(* Schneider Machine Expert - Basic project Projeto Charpy 3 - Prático V2, file version 3.0.0.0 *)
(* ProjectInformations: Name=Novo projeto *)

HARDWARE
  Cpu 0: TM221CE40R
  EthernetConfiguration: NetworkName=M221, IpAllocationMode=FixedAddress, IpAddress=10.0.0.20, SubnetMask=255.0.0.0
  SerialLineConfiguration: Baud=Baud19200, Parity=ParityEven, DataBits=DataBits8, StopBits=StopBits1, PhysicalMedium=PhysicalMediumRs485, TransmissionMode=TransmissionModeModbusRtu, SlaveId=1, Addressing=SlaveAddressing
  MastTask: UsePeriodScanMode=false, PeriodScan=100
  FastTask: Period=255
  CpuBehavior: StartingMode=StartAsPreviousState, AutoSaveRamOnEeprom=true, WatchdogPeriod=250

SYMBOLS  (address, symbol, comment, settings)
  %HSC0.V   VALOR_ENCODER  "Entrada de alta velocidade"
  %M0         "Engrenagem"
  %M1         "Motor Subir"
  %M2         "Motor Descer"
  %M3       LIB_CATRACA  "Solta Pêndulo"
  %M4       AUX_IMPACTO  "Subida do impacto"
  %M5         "Perdas"
  %M6       PERDAS_CONTAGEM  "Perdas_aux"
  %M7       PERDAS_SUBIR  "Aux_subir"
  %M8       ONOFF_ESTEIRA
  %M9       ESTEIRA  "Aux_Esteira"
  %M10      FALHA_PORTA  "Alerta de Falha"
  %M11      FALHA_SUBIDA  "Detecção de Falha"
  %M12      FALHA_DESCIDA  "Detecção de Falha"
  %M13      FALHA_MOTOR  "Alerta de Falha"
  %M14      FALHA_ÂNGULO
  %M15      M_SENSOR_PORTA  "Memória"
  %M16      M_SENSOR_BAIXO  "Memória"
  %M17      M_SENSOR_CIMA  "Memória"
  %M20        "ATRITO_OK"
  %M21        "ATRITO_FALHO"
  %M22      ATRITO_CONCLUIDO  "Fim do teste de atrito"
  %M23      ANG_0
  %M24      ANG_150
  %M25      AUX_ZERAR
  %M26      AUX_0
  %M27      AUX_150
  %M31      SENSOR_VIRTUAL_B  "Virtual_Baixo"
  %M32      SENSOR_VIRTUAL_C  "Virtual_Cima"
  %M100     ZERAR_SOFTWARE  "Botão de Zerar do Software"
  %M101     SUBIR_SOFTWARE  "Botão de Subir do Software"
  %M102     DESCER_SOFTWARE  "Botão de Descer do Software"
  %M103     IMPACTO_SOFTWARE  "Botão de Impacto do Software"
  %M105     PERDAS_SOFTWARE  "Botão de Perdas do Software"
  %S6       SB_TB1S  "Base de tempo de 1 s gerada por um relógio interno"
  %MW0      PULSOS_ENCODER  "Pulsos brutos do encoder"
  %MF2      ANGULO_ATUAL  "Ângulo instantâneo em Graus"
  %MF4      ANGULO_PICO  "Maior ângulo atingido no impacto"
  %MF6      ENERGIA_NOMINAL  "Capacidade da ponta do martelo"
  %MF8      ENERGIA_ABSORVIDA  "Resultado final do ensaio em Joules"
  %MF10     MF_10
  %MF12     MF_12
  %MF120    PERDAS_J  "Energia perdida por atrito em Joules"
  %TM0        [Preset=10, Base=OneSecond]
  %TM1        [Preset=15, Base=TenMilliSeconds]
  %TM2        [Preset=15, Base=TenMilliSeconds]
  %TM3        [Type=TP, Preset=1, Base=OneSecond]
  %TM5        "Zero 5s"  [Preset=5, Base=OneSecond]
  %TM6        "Zero 10s"  [Preset=10, Base=OneSecond]
  %I0.2     BOT_RESET  "Botão físico de zerar encoder e pico"
  %I0.10    SENSOR_PORTA  "Sensor se a porta está fechada"
  %I0.11    SENSOR_BAIXO  "Sensor se o braço está em baixo"
  %I0.12    SENSOR_CIMA  "Sensor se o braço está em cima"
  %I0.19    BOTÃO_ATRITO  "Botão que inicia o teste de atrito"
  %I0.20    BOTÃO_ZERAR  "Botão que zera a referência do encoder"
  %I0.21    BOTÃO_IMPACTO  "Botão que libera para o impacto"
  %I0.22    BOTÃO_DESCER  "Botão que aciona por 7s"
  %I0.23    BOTÃO_SUBIR  "Botão que aciona por 7s"
  %Q0.0     Q_0_0  "Encaixe Engrenagem"
  %Q0.1     Q_0_1  "Motor Subir"
  %Q0.2     Q_0_2  "Motor Descer"
  %Q0.3     Q_0_3  "Liberar Catraca"
  %Q0.4     Q_0_4  "Liga Esteira"
  %Q0.5     Q_0_5  "Led Porta"
  %Q0.14    Q_0_14
  %Q0.15    Q_0_15
  %IW0.0    IN_ANALOG  "Valor do Potenciômetro"  [Type=Type_0_10V, Scope=Scope_Normal, Minimum=0, Maximum=1000]
  %HSC0       [Type=CounterOrDownCounterBiPhasesX4, Preset=0, DedicatedInputs(DedicatedInput(Activated=true), DedicatedInput(Activated=true)), ReflexOutputs(ReflexOutput(Activated=false, LessThanS0=false, GreaterOrEqualThanS0=false, GreaterOrEqualThanS1=false), ReflexOutput(Activated=false, LessThanS0=false, GreaterOrEqualThanS0=false, GreaterOrEqualThanS1=false)), Thresholds(Threshold(ThresholdType=NotUsed, Pri]

POU Novo POU
  (* SectionNumber=1 *)

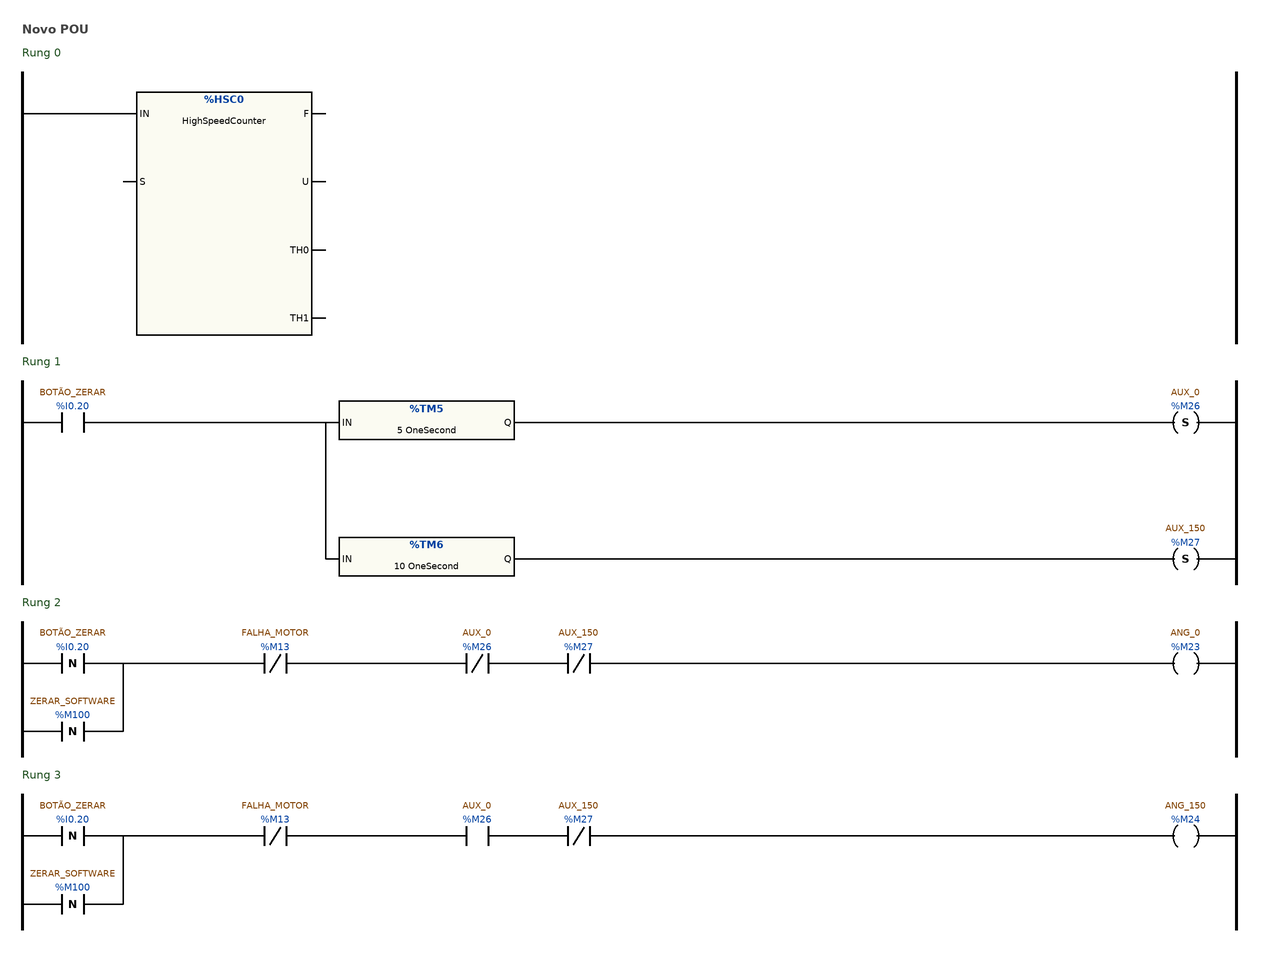

// Rung 0
  BLK %HSC0
  LD 1
  IN
  END_BLK
  // as ST:
  //   %HSC0(IN := TRUE);

// Rung 1
  LD 1
  MULTIFB
  LD 1
  AND %I0.20              (* BOTÃO_ZERAR *)
  ST %MW2009:X0
  BLK %TM5
  LD %MW2009:X0
  IN
  OUT_BLK
  LD Q
  S %M26                  (* AUX_0 *)
  END_BLK
  BLK %TM6
  LD %MW2009:X0
  IN
  OUT_BLK
  LD Q
  S %M27                  (* AUX_150 *)
  END_BLK
  MULTIFB
  // as ST:
  //   %TM5(IN := BOTÃO_ZERAR);
  //   IF %TM5.Q THEN AUX_0 := TRUE; END_IF;
  //   %TM6(IN := BOTÃO_ZERAR);
  //   IF %TM6.Q THEN AUX_150 := TRUE; END_IF;

// Rung 2
  LDF %I0.20              (* BOTÃO_ZERAR *)
  ORF %M100               (* ZERAR_SOFTWARE *)
  ANDN %M13               (* FALHA_MOTOR *)
  ANDN %M26               (* AUX_0 *)
  ANDN %M27               (* AUX_150 *)
  ST %M23                 (* ANG_0 *)
  // as ST:
  //   ANG_0 := (FALLING(BOTÃO_ZERAR) OR FALLING(ZERAR_SOFTWARE)) AND NOT FALHA_MOTOR AND NOT AUX_0 AND NOT AUX_150;

// Rung 3
  LDF %I0.20              (* BOTÃO_ZERAR *)
  ORF %M100               (* ZERAR_SOFTWARE *)
  ANDN %M13               (* FALHA_MOTOR *)
  AND %M26                (* AUX_0 *)
  ANDN %M27               (* AUX_150 *)
  ST %M24                 (* ANG_150 *)
  // as ST:
  //   ANG_150 := (FALLING(BOTÃO_ZERAR) OR FALLING(ZERAR_SOFTWARE)) AND NOT FALHA_MOTOR AND AUX_0 AND NOT AUX_150;

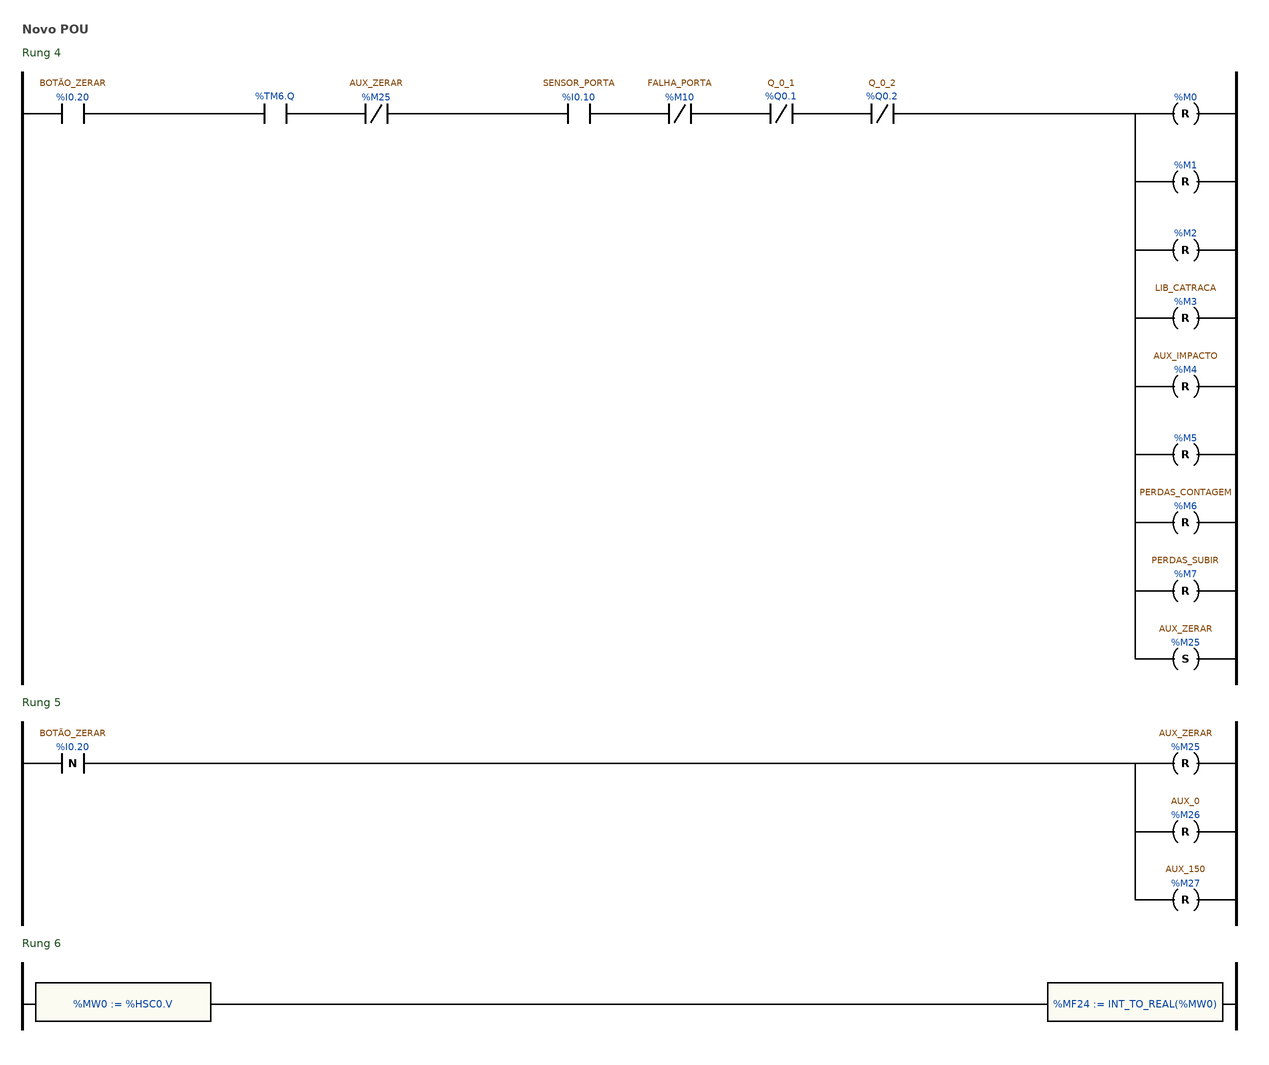

// Rung 4
  LD %I0.20               (* BOTÃO_ZERAR *)
  AND %TM6.Q
  ANDN %M25               (* AUX_ZERAR *)
  AND %I0.10              (* SENSOR_PORTA *)
  ANDN %M10               (* FALHA_PORTA *)
  ANDN %Q0.1              (* Q_0_1 *)
  ANDN %Q0.2              (* Q_0_2 *)
  R %M0
  R %M1
  R %M2
  R %M3                   (* LIB_CATRACA *)
  R %M4                   (* AUX_IMPACTO *)
  R %M5
  R %M6                   (* PERDAS_CONTAGEM *)
  R %M7                   (* PERDAS_SUBIR *)
  S %M25                  (* AUX_ZERAR *)
  // as ST:
  //   IF BOTÃO_ZERAR AND %TM6.Q AND NOT AUX_ZERAR AND SENSOR_PORTA AND NOT FALHA_PORTA AND NOT Q_0_1 AND NOT Q_0_2 THEN %M0 := FALSE; END_IF;
  //   IF BOTÃO_ZERAR AND %TM6.Q AND NOT AUX_ZERAR AND SENSOR_PORTA AND NOT FALHA_PORTA AND NOT Q_0_1 AND NOT Q_0_2 THEN %M1 := FALSE; END_IF;
  //   IF BOTÃO_ZERAR AND %TM6.Q AND NOT AUX_ZERAR AND SENSOR_PORTA AND NOT FALHA_PORTA AND NOT Q_0_1 AND NOT Q_0_2 THEN %M2 := FALSE; END_IF;
  //   IF BOTÃO_ZERAR AND %TM6.Q AND NOT AUX_ZERAR AND SENSOR_PORTA AND NOT FALHA_PORTA AND NOT Q_0_1 AND NOT Q_0_2 THEN LIB_CATRACA := FALSE; END_IF;
  //   IF BOTÃO_ZERAR AND %TM6.Q AND NOT AUX_ZERAR AND SENSOR_PORTA AND NOT FALHA_PORTA AND NOT Q_0_1 AND NOT Q_0_2 THEN AUX_IMPACTO := FALSE; END_IF;
  //   IF BOTÃO_ZERAR AND %TM6.Q AND NOT AUX_ZERAR AND SENSOR_PORTA AND NOT FALHA_PORTA AND NOT Q_0_1 AND NOT Q_0_2 THEN %M5 := FALSE; END_IF;
  //   IF BOTÃO_ZERAR AND %TM6.Q AND NOT AUX_ZERAR AND SENSOR_PORTA AND NOT FALHA_PORTA AND NOT Q_0_1 AND NOT Q_0_2 THEN PERDAS_CONTAGEM := FALSE; END_IF;
  //   IF BOTÃO_ZERAR AND %TM6.Q AND NOT AUX_ZERAR AND SENSOR_PORTA AND NOT FALHA_PORTA AND NOT Q_0_1 AND NOT Q_0_2 THEN PERDAS_SUBIR := FALSE; END_IF;
  //   IF BOTÃO_ZERAR AND %TM6.Q AND NOT AUX_ZERAR AND SENSOR_PORTA AND NOT FALHA_PORTA AND NOT Q_0_1 AND NOT Q_0_2 THEN AUX_ZERAR := TRUE; END_IF;

// Rung 5
  LDF %I0.20              (* BOTÃO_ZERAR *)
  R %M25                  (* AUX_ZERAR *)
  R %M26                  (* AUX_0 *)
  R %M27                  (* AUX_150 *)
  // as ST:
  //   IF FALLING(BOTÃO_ZERAR) THEN AUX_ZERAR := FALSE; END_IF;
  //   IF FALLING(BOTÃO_ZERAR) THEN AUX_0 := FALSE; END_IF;
  //   IF FALLING(BOTÃO_ZERAR) THEN AUX_150 := FALSE; END_IF;

// Rung 6
  LD 1
  OPER [ %MW0 := %HSC0.V ](* PULSOS_ENCODER *)
  [ %MF24 := INT_TO_REAL ( %MW0 ) ](* PULSOS_ENCODER *)
  // as ST:
  //   PULSOS_ENCODER := %HSC0.V;
  //   %MF24 := INT_TO_REAL ( PULSOS_ENCODER );

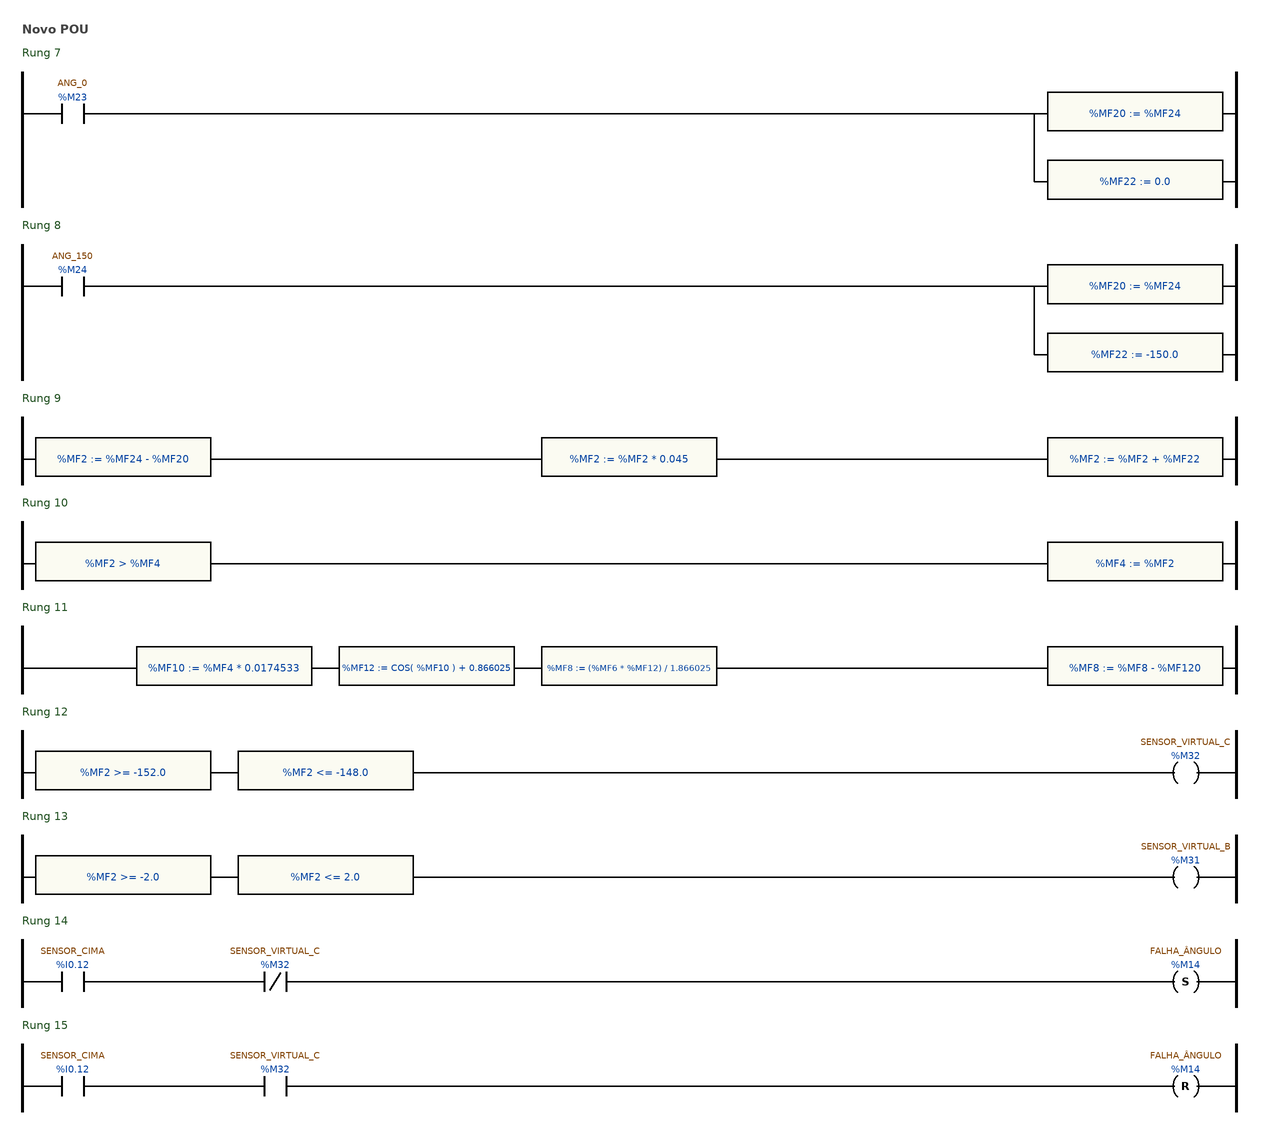

// Rung 7
  LD %M23                 (* ANG_0 *)
  [ %MF20 := %MF24 ]
  [ %MF22 := 0.0 ]
  // as ST:
  //   IF ANG_0 THEN %MF20 := %MF24; END_IF;
  //   IF ANG_0 THEN %MF22 := 0.0; END_IF;

// Rung 8
  LD %M24                 (* ANG_150 *)
  [ %MF20 := %MF24 ]
  [ %MF22 := -150.0 ]
  // as ST:
  //   IF ANG_150 THEN %MF20 := %MF24; END_IF;
  //   IF ANG_150 THEN %MF22 := -150.0; END_IF;

// Rung 9
  LD 1
  OPER [ %MF2 := %MF24 - %MF20 ](* ANGULO_ATUAL *)
  OPER [ %MF2 := %MF2 * 0.045 ](* ANGULO_ATUAL, ANGULO_ATUAL *)
  [ %MF2 := %MF2 + %MF22 ](* ANGULO_ATUAL, ANGULO_ATUAL *)
  // as ST:
  //   ANGULO_ATUAL := %MF24 - %MF20;
  //   ANGULO_ATUAL := ANGULO_ATUAL * 0.045;
  //   ANGULO_ATUAL := ANGULO_ATUAL + %MF22;

// Rung 10
  LD [ %MF2 > %MF4 ]      (* ANGULO_ATUAL, ANGULO_PICO *)
  [ %MF4 := %MF2 ]        (* ANGULO_PICO, ANGULO_ATUAL *)
  // as ST:
  //   IF ANGULO_ATUAL > ANGULO_PICO THEN ANGULO_PICO := ANGULO_ATUAL; END_IF;

// Rung 11
  LD 1
  OPER [ %MF10 := %MF4 * 0.0174533 ](* MF_10, ANGULO_PICO *)
  OPER [%MF12 := COS( %MF10 ) + 0.866025](* MF_12, MF_10 *)
  OPER [%MF8 := (%MF6 * %MF12) / 1.866025](* ENERGIA_ABSORVIDA, ENERGIA_NOMINAL, MF_12 *)
  [ %MF8 := %MF8 - %MF120 ](* ENERGIA_ABSORVIDA, ENERGIA_ABSORVIDA, PERDAS_J *)
  // as ST:
  //   MF_10 := ANGULO_PICO * 0.0174533;
  //   MF_12 := COS( MF_10 ) + 0.866025;
  //   ENERGIA_ABSORVIDA := (ENERGIA_NOMINAL * MF_12) / 1.866025;
  //   ENERGIA_ABSORVIDA := ENERGIA_ABSORVIDA - PERDAS_J;

// Rung 12
  LD [ %MF2 >= -152.0 ]   (* ANGULO_ATUAL *)
  AND [ %MF2 <= -148.0 ]  (* ANGULO_ATUAL *)
  ST %M32                 (* SENSOR_VIRTUAL_C *)
  // as ST:
  //   SENSOR_VIRTUAL_C := ANGULO_ATUAL >= -152.0 AND ANGULO_ATUAL <= -148.0;

// Rung 13
  LD [ %MF2 >= -2.0 ]     (* ANGULO_ATUAL *)
  AND [ %MF2 <= 2.0 ]     (* ANGULO_ATUAL *)
  ST %M31                 (* SENSOR_VIRTUAL_B *)
  // as ST:
  //   SENSOR_VIRTUAL_B := ANGULO_ATUAL >= -2.0 AND ANGULO_ATUAL <= 2.0;

// Rung 14
  LD %I0.12               (* SENSOR_CIMA *)
  ANDN %M32               (* SENSOR_VIRTUAL_C *)
  S %M14                  (* FALHA_ÂNGULO *)
  // as ST:
  //   IF SENSOR_CIMA AND NOT SENSOR_VIRTUAL_C THEN FALHA_ÂNGULO := TRUE; END_IF;

// Rung 15
  LD %I0.12               (* SENSOR_CIMA *)
  AND %M32                (* SENSOR_VIRTUAL_C *)
  R %M14                  (* FALHA_ÂNGULO *)
  // as ST:
  //   IF SENSOR_CIMA AND SENSOR_VIRTUAL_C THEN FALHA_ÂNGULO := FALSE; END_IF;

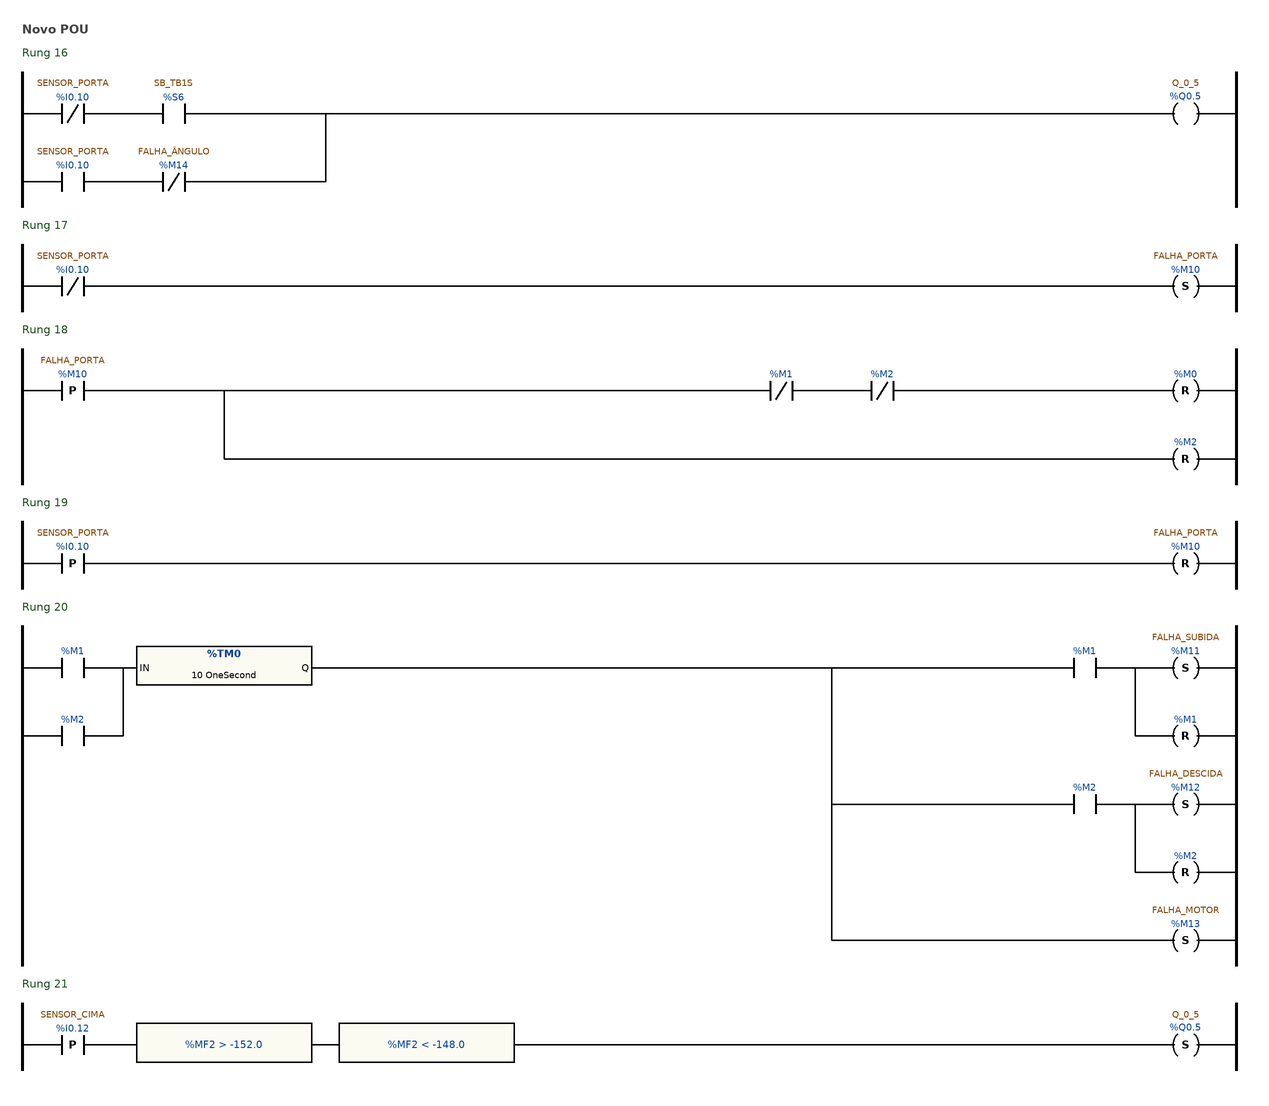

// Rung 16
  LDN %I0.10              (* SENSOR_PORTA *)
  AND %S6                 (* SB_TB1S *)
  OR( %I0.10              (* SENSOR_PORTA *)
  ANDN %M14               (* FALHA_ÂNGULO *)
  )
  ST %Q0.5                (* Q_0_5 *)
  // as ST:
  //   Q_0_5 := NOT SENSOR_PORTA AND SB_TB1S OR SENSOR_PORTA AND NOT FALHA_ÂNGULO;

// Rung 17
  LDN %I0.10              (* SENSOR_PORTA *)
  S %M10                  (* FALHA_PORTA *)
  // as ST:
  //   IF NOT SENSOR_PORTA THEN FALHA_PORTA := TRUE; END_IF;

// Rung 18
  LDR %M10                (* FALHA_PORTA *)
  MPS
  ANDN %M1
  ANDN %M2
  R %M0
  MPP
  R %M2
  // as ST:
  //   IF RISING(FALHA_PORTA) AND NOT %M1 AND NOT %M2 THEN %M0 := FALSE; END_IF;
  //   IF RISING(FALHA_PORTA) THEN %M2 := FALSE; END_IF;

// Rung 19
  LDR %I0.10              (* SENSOR_PORTA *)
  R %M10                  (* FALHA_PORTA *)
  // as ST:
  //   IF RISING(SENSOR_PORTA) THEN FALHA_PORTA := FALSE; END_IF;

// Rung 20
  BLK %TM0
  LD %M1
  OR %M2
  IN
  OUT_BLK
  LD Q
  MPS
  AND %M1
  S %M11                  (* FALHA_SUBIDA *)
  R %M1
  MRD
  AND %M2
  S %M12                  (* FALHA_DESCIDA *)
  R %M2
  MPP
  S %M13                  (* FALHA_MOTOR *)
  END_BLK
  // as ST:
  //   %TM0(IN := %M1 OR %M2);
  //   IF %TM0.Q AND %M1 THEN FALHA_SUBIDA := TRUE; END_IF;
  //   IF %TM0.Q AND %M1 THEN %M1 := FALSE; END_IF;
  //   IF %TM0.Q AND %M2 THEN FALHA_DESCIDA := TRUE; END_IF;
  //   IF %TM0.Q AND %M2 THEN %M2 := FALSE; END_IF;
  //   IF %TM0.Q THEN FALHA_MOTOR := TRUE; END_IF;

// Rung 21
  LDR %I0.12              (* SENSOR_CIMA *)
  AND [ %MF2 > -152.0 ]   (* ANGULO_ATUAL *)
  AND [ %MF2 < -148.0 ]   (* ANGULO_ATUAL *)
  S %Q0.5                 (* Q_0_5 *)
  // as ST:
  //   IF RISING(SENSOR_CIMA) AND ANGULO_ATUAL > -152.0 AND ANGULO_ATUAL < -148.0 THEN Q_0_5 := TRUE; END_IF;

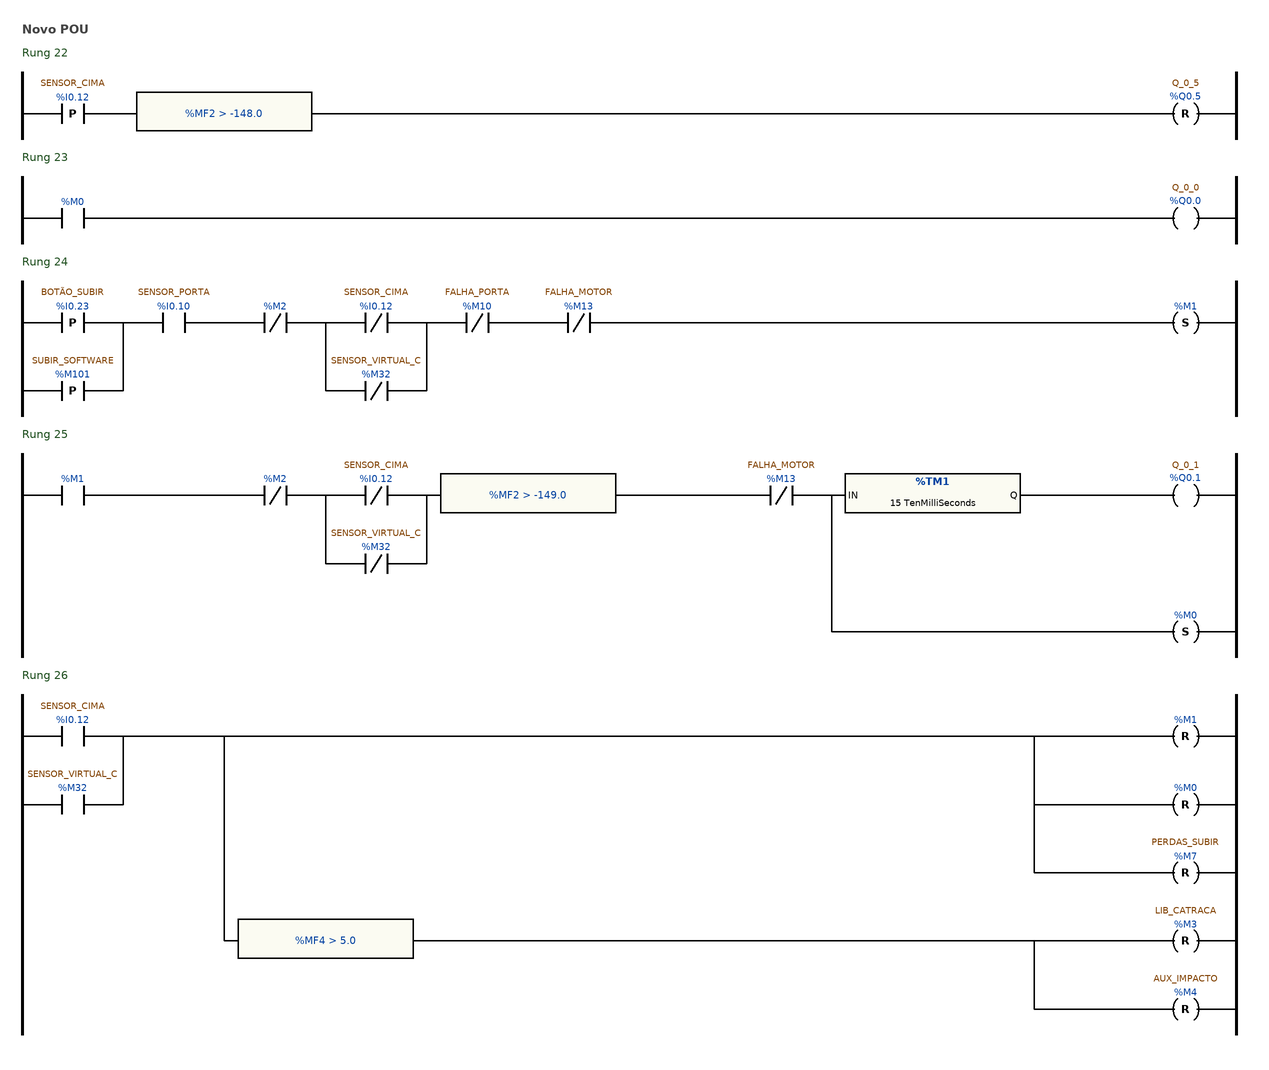

// Rung 22
  LDR %I0.12              (* SENSOR_CIMA *)
  AND [ %MF2 > -148.0 ]   (* ANGULO_ATUAL *)
  R %Q0.5                 (* Q_0_5 *)
  // as ST:
  //   IF RISING(SENSOR_CIMA) AND ANGULO_ATUAL > -148.0 THEN Q_0_5 := FALSE; END_IF;

// Rung 23
  LD %M0
  ST %Q0.0                (* Q_0_0 *)
  // as ST:
  //   Q_0_0 := %M0;

// Rung 24
  LDR %I0.23              (* BOTÃO_SUBIR *)
  ORR %M101               (* SUBIR_SOFTWARE *)
  AND %I0.10              (* SENSOR_PORTA *)
  ANDN %M2
  AND(N %I0.12            (* SENSOR_CIMA *)
  ORN %M32                (* SENSOR_VIRTUAL_C *)
  )
  ANDN %M10               (* FALHA_PORTA *)
  ANDN %M13               (* FALHA_MOTOR *)
  S %M1
  // as ST:
  //   IF (RISING(BOTÃO_SUBIR) OR RISING(SUBIR_SOFTWARE)) AND SENSOR_PORTA AND NOT %M2 AND (NOT SENSOR_CIMA OR NOT SENSOR_VIRTUAL_C) AND NOT FALHA_PORTA AND NOT FALHA_MOTOR THEN %M1 := TRUE; END_IF;

// Rung 25
  LD 1
  MULTIFB
  LD 1
  AND %M1
  ANDN %M2
  AND(N %I0.12            (* SENSOR_CIMA *)
  ORN %M32                (* SENSOR_VIRTUAL_C *)
  )
  AND [ %MF2 > -149.0 ]   (* ANGULO_ATUAL *)
  ANDN %M13               (* FALHA_MOTOR *)
  ST %MW2009:X0
  BLK %TM1
  LD %MW2009:X0
  IN
  OUT_BLK
  LD Q
  ST %Q0.1                (* Q_0_1 *)
  END_BLK
  LD %MW2009:X0
  S %M0
  MULTIFB
  // as ST:
  //   %TM1(IN := %M1 AND NOT %M2 AND (NOT SENSOR_CIMA OR NOT SENSOR_VIRTUAL_C) AND ANGULO_ATUAL > -149.0 AND NOT FALHA_MOTOR);
  //   Q_0_1 := %TM1.Q;
  //   IF %M1 AND NOT %M2 AND (NOT SENSOR_CIMA OR NOT SENSOR_VIRTUAL_C) AND ANGULO_ATUAL > -149.0 AND NOT FALHA_MOTOR THEN %M0 := TRUE; END_IF;

// Rung 26
  LD %I0.12               (* SENSOR_CIMA *)
  OR %M32                 (* SENSOR_VIRTUAL_C *)
  MPS
  R %M1
  R %M0
  R %M7                   (* PERDAS_SUBIR *)
  MPP
  AND [ %MF4 > 5.0 ]      (* ANGULO_PICO *)
  R %M3                   (* LIB_CATRACA *)
  R %M4                   (* AUX_IMPACTO *)
  // as ST:
  //   IF SENSOR_CIMA OR SENSOR_VIRTUAL_C THEN %M1 := FALSE; END_IF;
  //   IF SENSOR_CIMA OR SENSOR_VIRTUAL_C THEN %M0 := FALSE; END_IF;
  //   IF SENSOR_CIMA OR SENSOR_VIRTUAL_C THEN PERDAS_SUBIR := FALSE; END_IF;
  //   IF (SENSOR_CIMA OR SENSOR_VIRTUAL_C) AND ANGULO_PICO > 5.0 THEN LIB_CATRACA := FALSE; END_IF;
  //   IF (SENSOR_CIMA OR SENSOR_VIRTUAL_C) AND ANGULO_PICO > 5.0 THEN AUX_IMPACTO := FALSE; END_IF;

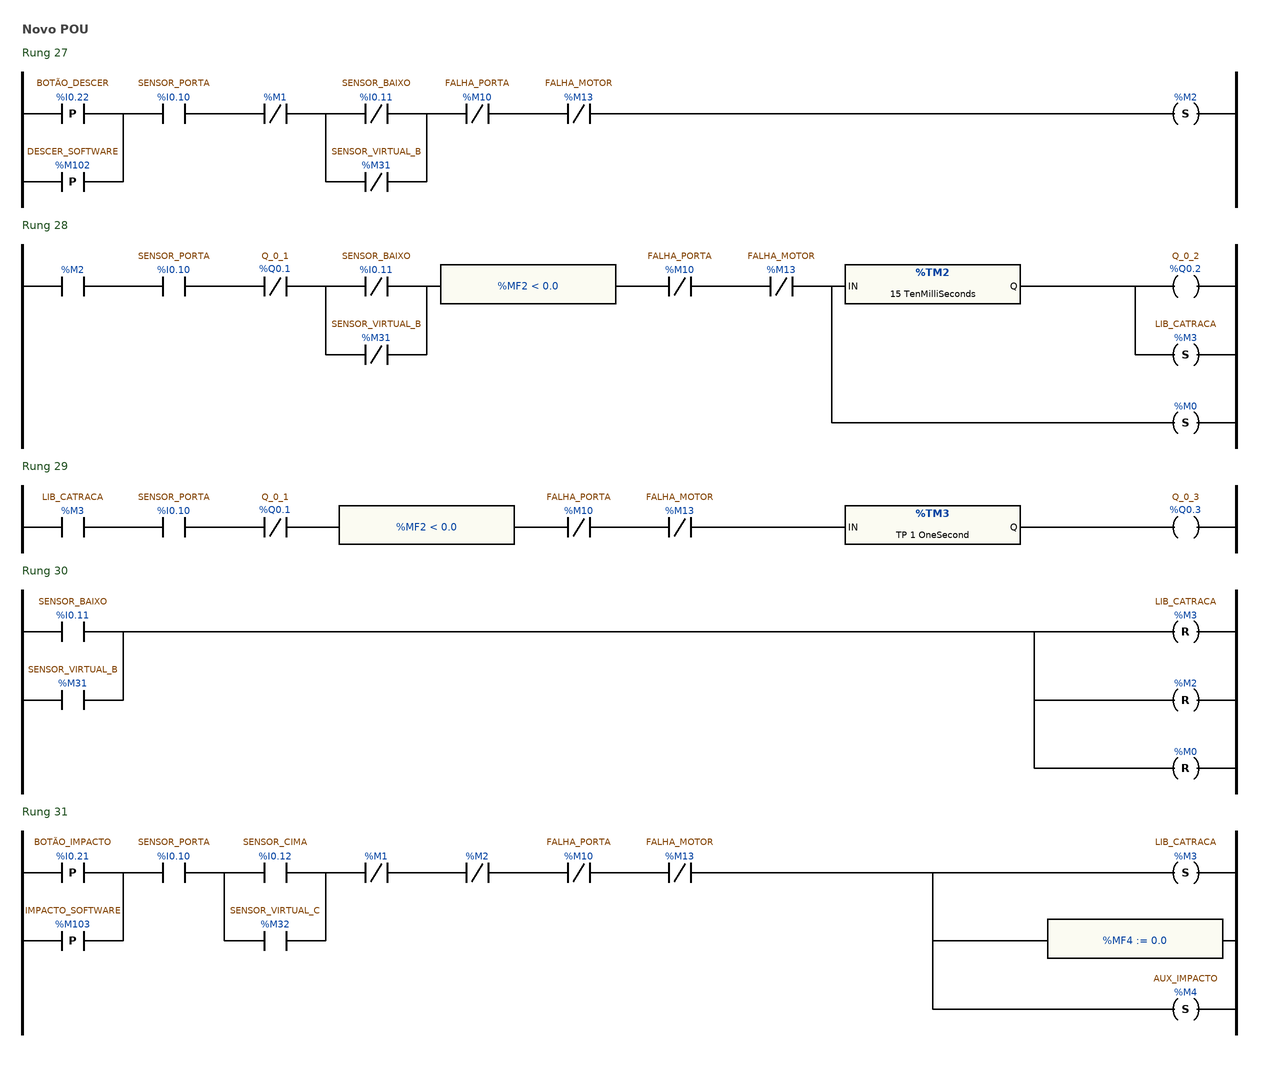

// Rung 27
  LDR %I0.22              (* BOTÃO_DESCER *)
  ORR %M102               (* DESCER_SOFTWARE *)
  AND %I0.10              (* SENSOR_PORTA *)
  ANDN %M1
  AND(N %I0.11            (* SENSOR_BAIXO *)
  ORN %M31                (* SENSOR_VIRTUAL_B *)
  )
  ANDN %M10               (* FALHA_PORTA *)
  ANDN %M13               (* FALHA_MOTOR *)
  S %M2
  // as ST:
  //   IF (RISING(BOTÃO_DESCER) OR RISING(DESCER_SOFTWARE)) AND SENSOR_PORTA AND NOT %M1 AND (NOT SENSOR_BAIXO OR NOT SENSOR_VIRTUAL_B) AND NOT FALHA_PORTA AND NOT FALHA_MOTOR THEN %M2 := TRUE; END_IF;

// Rung 28
  LD 1
  MULTIFB
  LD 1
  AND %M2
  AND %I0.10              (* SENSOR_PORTA *)
  ANDN %Q0.1              (* Q_0_1 *)
  AND(N %I0.11            (* SENSOR_BAIXO *)
  ORN %M31                (* SENSOR_VIRTUAL_B *)
  )
  AND [ %MF2 < 0.0 ]      (* ANGULO_ATUAL *)
  ANDN %M10               (* FALHA_PORTA *)
  ANDN %M13               (* FALHA_MOTOR *)
  ST %MW2009:X0
  BLK %TM2
  LD %MW2009:X0
  IN
  OUT_BLK
  LD Q
  ST %Q0.2                (* Q_0_2 *)
  S %M3                   (* LIB_CATRACA *)
  END_BLK
  LD %MW2009:X0
  S %M0
  MULTIFB
  // as ST:
  //   %TM2(IN := %M2 AND SENSOR_PORTA AND NOT Q_0_1 AND (NOT SENSOR_BAIXO OR NOT SENSOR_VIRTUAL_B) AND ANGULO_ATUAL < 0.0 AND NOT FALHA_PORTA AND NOT FALHA_MOTOR);
  //   Q_0_2 := %TM2.Q;
  //   IF %TM2.Q THEN LIB_CATRACA := TRUE; END_IF;
  //   IF %M2 AND SENSOR_PORTA AND NOT Q_0_1 AND (NOT SENSOR_BAIXO OR NOT SENSOR_VIRTUAL_B) AND ANGULO_ATUAL < 0.0 AND NOT FALHA_PORTA AND NOT FALHA_MOTOR THEN %M0 := TRUE; END_IF;

// Rung 29
  BLK %TM3
  LD %M3                  (* LIB_CATRACA *)
  AND %I0.10              (* SENSOR_PORTA *)
  ANDN %Q0.1              (* Q_0_1 *)
  AND [ %MF2 < 0.0 ]      (* ANGULO_ATUAL *)
  ANDN %M10               (* FALHA_PORTA *)
  ANDN %M13               (* FALHA_MOTOR *)
  IN
  OUT_BLK
  LD Q
  ST %Q0.3                (* Q_0_3 *)
  END_BLK
  // as ST:
  //   %TM3(IN := LIB_CATRACA AND SENSOR_PORTA AND NOT Q_0_1 AND ANGULO_ATUAL < 0.0 AND NOT FALHA_PORTA AND NOT FALHA_MOTOR);
  //   Q_0_3 := %TM3.Q;

// Rung 30
  LD %I0.11               (* SENSOR_BAIXO *)
  OR %M31                 (* SENSOR_VIRTUAL_B *)
  R %M3                   (* LIB_CATRACA *)
  R %M2
  R %M0
  // as ST:
  //   IF SENSOR_BAIXO OR SENSOR_VIRTUAL_B THEN LIB_CATRACA := FALSE; END_IF;
  //   IF SENSOR_BAIXO OR SENSOR_VIRTUAL_B THEN %M2 := FALSE; END_IF;
  //   IF SENSOR_BAIXO OR SENSOR_VIRTUAL_B THEN %M0 := FALSE; END_IF;

// Rung 31
  LDR %I0.21              (* BOTÃO_IMPACTO *)
  ORR %M103               (* IMPACTO_SOFTWARE *)
  AND %I0.10              (* SENSOR_PORTA *)
  AND( %I0.12             (* SENSOR_CIMA *)
  OR %M32                 (* SENSOR_VIRTUAL_C *)
  )
  ANDN %M1
  ANDN %M2
  ANDN %M10               (* FALHA_PORTA *)
  ANDN %M13               (* FALHA_MOTOR *)
  S %M3                   (* LIB_CATRACA *)
  [ %MF4 := 0.0 ]         (* ANGULO_PICO *)
  S %M4                   (* AUX_IMPACTO *)
  // as ST:
  //   IF (RISING(BOTÃO_IMPACTO) OR RISING(IMPACTO_SOFTWARE)) AND SENSOR_PORTA AND (SENSOR_CIMA OR SENSOR_VIRTUAL_C) AND NOT %M1 AND NOT %M2 AND NOT FALHA_PORTA AND NOT FALHA_MOTOR THEN LIB_CATRACA := TRUE; END_IF;
  //   IF (RISING(BOTÃO_IMPACTO) OR RISING(IMPACTO_SOFTWARE)) AND SENSOR_PORTA AND (SENSOR_CIMA OR SENSOR_VIRTUAL_C) AND NOT %M1 AND NOT %M2 AND NOT FALHA_PORTA AND NOT FALHA_MOTOR THEN ANGULO_PICO := 0.0; END_IF;
  //   IF (RISING(BOTÃO_IMPACTO) OR RISING(IMPACTO_SOFTWARE)) AND SENSOR_PORTA AND (SENSOR_CIMA OR SENSOR_VIRTUAL_C) AND NOT %M1 AND NOT %M2 AND NOT FALHA_PORTA AND NOT FALHA_MOTOR THEN AUX_IMPACTO := TRUE; END_IF;

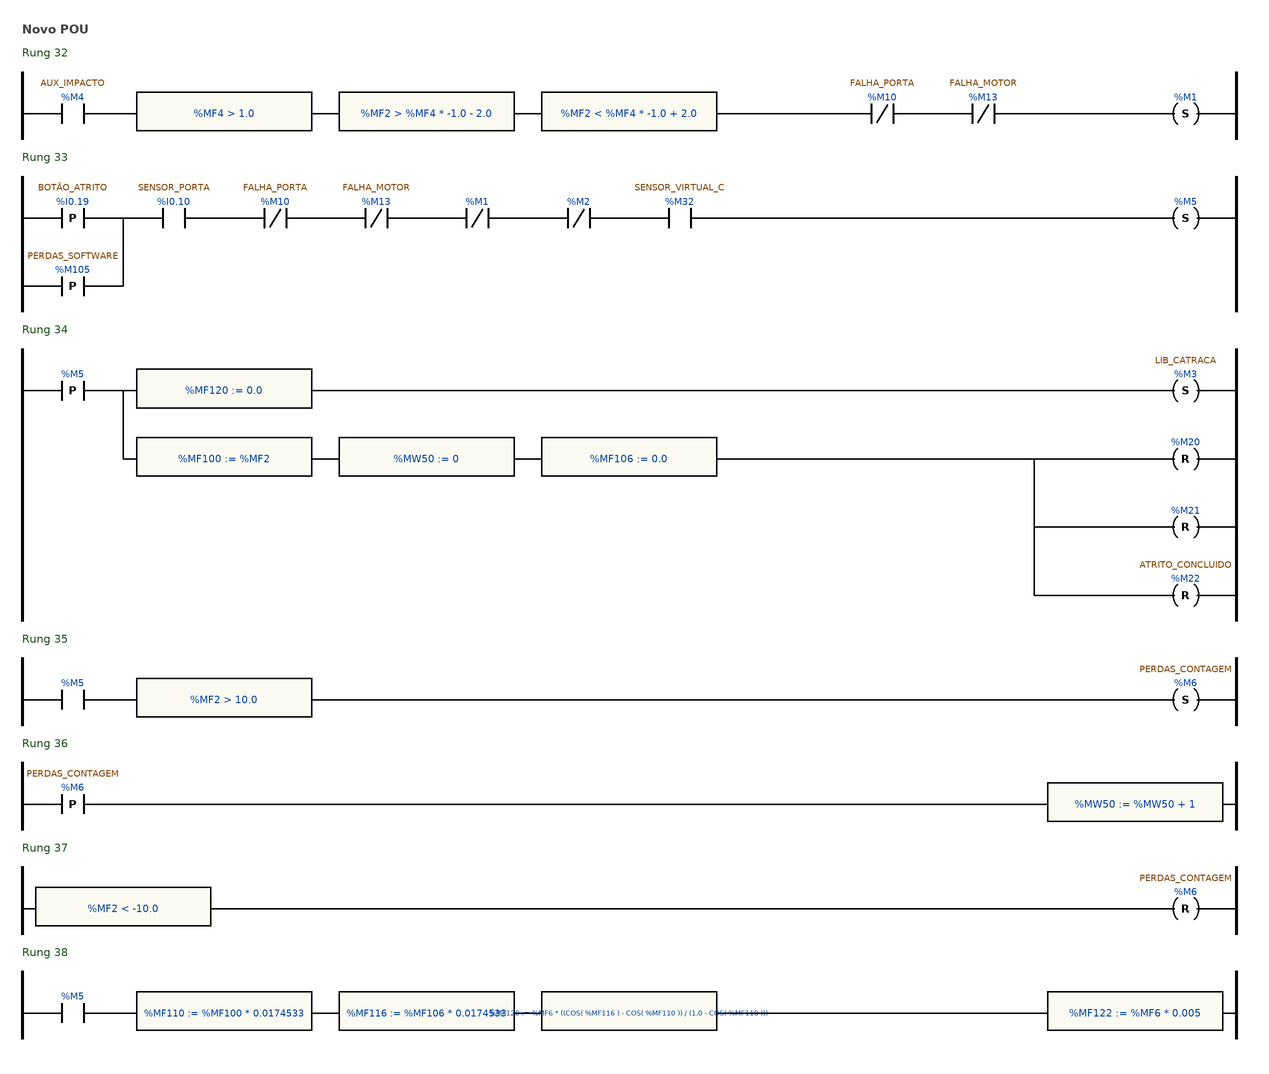

// Rung 32
  LD %M4                  (* AUX_IMPACTO *)
  AND [ %MF4 > 1.0 ]      (* ANGULO_PICO *)
  AND [%MF2 > %MF4 * -1.0 - 2.0](* ANGULO_ATUAL, ANGULO_PICO *)
  AND [%MF2 < %MF4 * -1.0 + 2.0](* ANGULO_ATUAL, ANGULO_PICO *)
  ANDN %M10               (* FALHA_PORTA *)
  ANDN %M13               (* FALHA_MOTOR *)
  S %M1
  // as ST:
  //   IF AUX_IMPACTO AND ANGULO_PICO > 1.0 AND ANGULO_ATUAL > ANGULO_PICO * -1.0 - 2.0 AND ANGULO_ATUAL < ANGULO_PICO * -1.0 + 2.0 AND NOT FALHA_PORTA AND NOT FALHA_MOTOR THEN %M1 := TRUE; END_IF;

// Rung 33
  LDR %I0.19              (* BOTÃO_ATRITO *)
  ORR %M105               (* PERDAS_SOFTWARE *)
  AND %I0.10              (* SENSOR_PORTA *)
  ANDN %M10               (* FALHA_PORTA *)
  ANDN %M13               (* FALHA_MOTOR *)
  ANDN %M1
  ANDN %M2
  AND %M32                (* SENSOR_VIRTUAL_C *)
  S %M5
  // as ST:
  //   IF (RISING(BOTÃO_ATRITO) OR RISING(PERDAS_SOFTWARE)) AND SENSOR_PORTA AND NOT FALHA_PORTA AND NOT FALHA_MOTOR AND NOT %M1 AND NOT %M2 AND SENSOR_VIRTUAL_C THEN %M5 := TRUE; END_IF;

// Rung 34
  LDR %M5
  MPS
  OPER [ %MF120 := 0.0 ]  (* PERDAS_J *)
  S %M3                   (* LIB_CATRACA *)
  MPP
  OPER [ %MF100 := %MF2 ] (* ANGULO_ATUAL *)
  OPER [ %MW50 := 0 ]
  OPER [ %MF106 := 0.0 ]
  R %M20
  R %M21
  R %M22                  (* ATRITO_CONCLUIDO *)
  // as ST:
  //   IF RISING(%M5) THEN PERDAS_J := 0.0; END_IF;
  //   IF RISING(%M5) THEN LIB_CATRACA := TRUE; END_IF;
  //   IF RISING(%M5) THEN %MF100 := ANGULO_ATUAL; END_IF;
  //   IF RISING(%M5) THEN %MW50 := 0; END_IF;
  //   IF RISING(%M5) THEN %MF106 := 0.0; END_IF;
  //   IF RISING(%M5) THEN %M20 := FALSE; END_IF;
  //   IF RISING(%M5) THEN %M21 := FALSE; END_IF;
  //   IF RISING(%M5) THEN ATRITO_CONCLUIDO := FALSE; END_IF;

// Rung 35
  LD %M5
  AND [ %MF2 > 10.0 ]     (* ANGULO_ATUAL *)
  S %M6                   (* PERDAS_CONTAGEM *)
  // as ST:
  //   IF %M5 AND ANGULO_ATUAL > 10.0 THEN PERDAS_CONTAGEM := TRUE; END_IF;

// Rung 36
  LDR %M6                 (* PERDAS_CONTAGEM *)
  [ %MW50 := %MW50 + 1 ]
  // as ST:
  //   IF RISING(PERDAS_CONTAGEM) THEN %MW50 := %MW50 + 1; END_IF;

// Rung 37
  LD [ %MF2 < -10.0 ]     (* ANGULO_ATUAL *)
  R %M6                   (* PERDAS_CONTAGEM *)
  // as ST:
  //   IF ANGULO_ATUAL < -10.0 THEN PERDAS_CONTAGEM := FALSE; END_IF;

// Rung 38
  LD %M5
  OPER [ %MF110 := %MF100 * 0.0174533 ]
  OPER [ %MF116 := %MF106 * 0.0174533 ]
  OPER [%MF120 := %MF6 * ((COS( %MF116 ) - COS( %MF110 )) / (1.0 - COS( %MF110 )))](* PERDAS_J, ENERGIA_NOMINAL *)
  [ %MF122 := %MF6 * 0.005 ](* ENERGIA_NOMINAL *)
  // as ST:
  //   IF %M5 THEN %MF110 := %MF100 * 0.0174533; END_IF;
  //   IF %M5 THEN %MF116 := %MF106 * 0.0174533; END_IF;
  //   IF %M5 THEN PERDAS_J := ENERGIA_NOMINAL * ((COS( %MF116 ) - COS( %MF110 )) / (1.0 - COS( %MF110 ))); END_IF;
  //   IF %M5 THEN %MF122 := ENERGIA_NOMINAL * 0.005; END_IF;

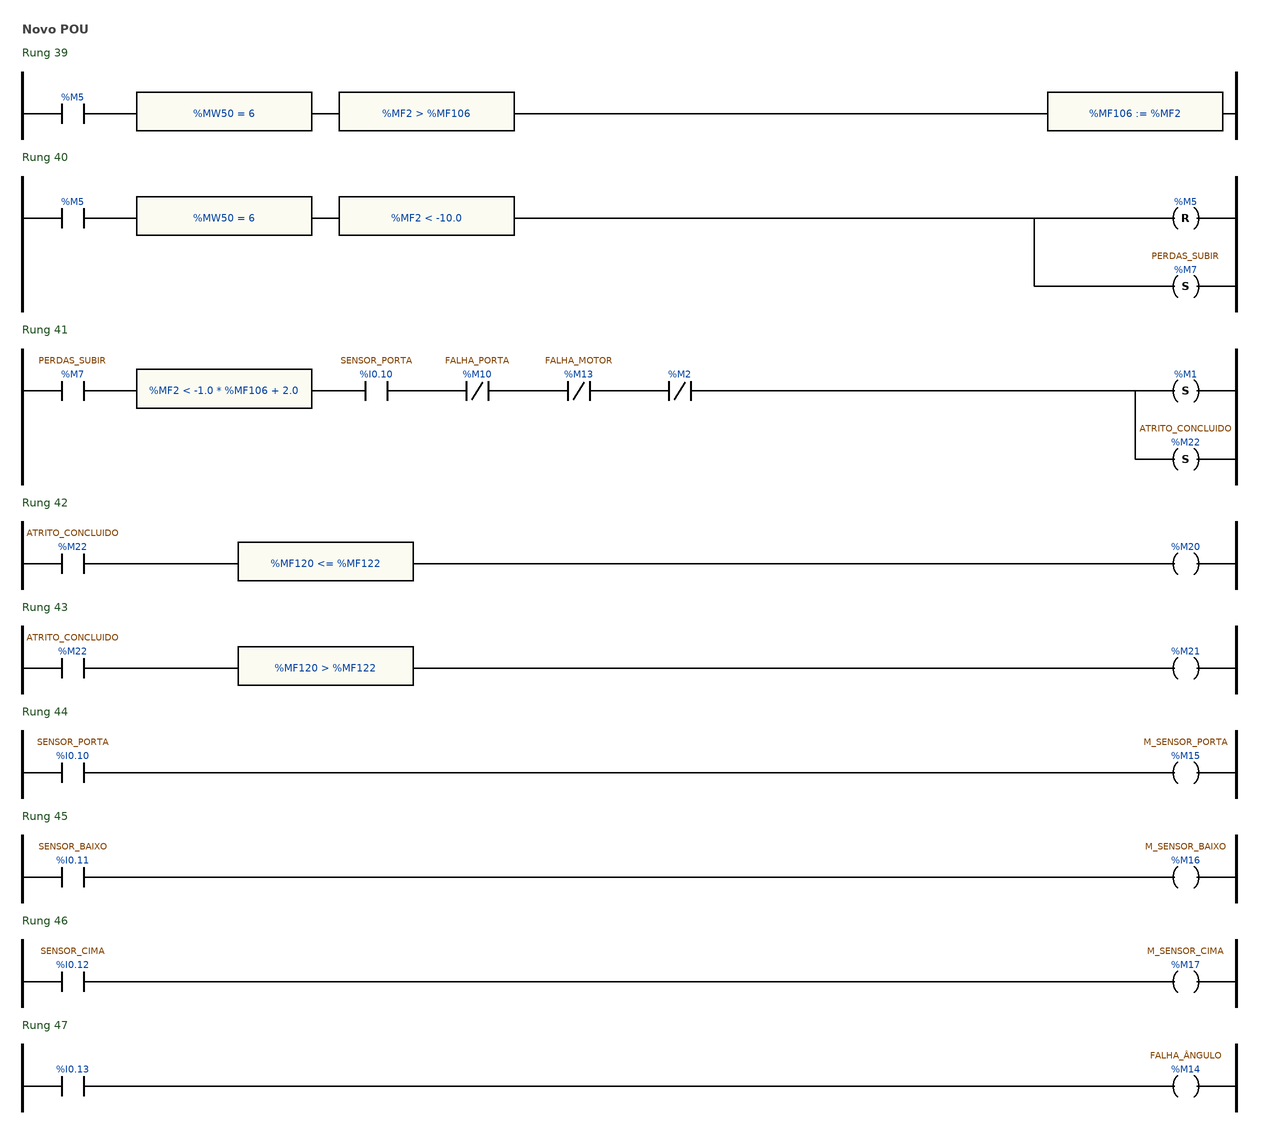

// Rung 39
  LD %M5
  AND [ %MW50 = 6 ]
  AND [ %MF2 > %MF106 ]   (* ANGULO_ATUAL *)
  [ %MF106 := %MF2 ]      (* ANGULO_ATUAL *)
  // as ST:
  //   IF %M5 AND %MW50 = 6 AND ANGULO_ATUAL > %MF106 THEN %MF106 := ANGULO_ATUAL; END_IF;

// Rung 40
  LD %M5
  AND [ %MW50 = 6 ]
  AND [ %MF2 < -10.0 ]    (* ANGULO_ATUAL *)
  R %M5
  S %M7                   (* PERDAS_SUBIR *)
  // as ST:
  //   _t1 := %M5 AND %MW50 = 6 AND ANGULO_ATUAL < -10.0;
  //   IF _t1 THEN %M5 := FALSE; END_IF;
  //   IF _t1 THEN PERDAS_SUBIR := TRUE; END_IF;

// Rung 41
  LD %M7                  (* PERDAS_SUBIR *)
  AND [%MF2 < -1.0 * %MF106 + 2.0](* ANGULO_ATUAL *)
  AND %I0.10              (* SENSOR_PORTA *)
  ANDN %M10               (* FALHA_PORTA *)
  ANDN %M13               (* FALHA_MOTOR *)
  ANDN %M2
  S %M1
  S %M22                  (* ATRITO_CONCLUIDO *)
  // as ST:
  //   IF PERDAS_SUBIR AND ANGULO_ATUAL < -1.0 * %MF106 + 2.0 AND SENSOR_PORTA AND NOT FALHA_PORTA AND NOT FALHA_MOTOR AND NOT %M2 THEN %M1 := TRUE; END_IF;
  //   IF PERDAS_SUBIR AND ANGULO_ATUAL < -1.0 * %MF106 + 2.0 AND SENSOR_PORTA AND NOT FALHA_PORTA AND NOT FALHA_MOTOR AND NOT %M2 THEN ATRITO_CONCLUIDO := TRUE; END_IF;

// Rung 42
  LD %M22                 (* ATRITO_CONCLUIDO *)
  AND [ %MF120 <= %MF122 ](* PERDAS_J *)
  ST %M20
  // as ST:
  //   %M20 := ATRITO_CONCLUIDO AND PERDAS_J <= %MF122;

// Rung 43
  LD %M22                 (* ATRITO_CONCLUIDO *)
  AND [ %MF120 > %MF122 ] (* PERDAS_J *)
  ST %M21
  // as ST:
  //   %M21 := ATRITO_CONCLUIDO AND PERDAS_J > %MF122;

// Rung 44
  LD %I0.10               (* SENSOR_PORTA *)
  ST %M15                 (* M_SENSOR_PORTA *)
  // as ST:
  //   M_SENSOR_PORTA := SENSOR_PORTA;

// Rung 45
  LD %I0.11               (* SENSOR_BAIXO *)
  ST %M16                 (* M_SENSOR_BAIXO *)
  // as ST:
  //   M_SENSOR_BAIXO := SENSOR_BAIXO;

// Rung 46
  LD %I0.12               (* SENSOR_CIMA *)
  ST %M17                 (* M_SENSOR_CIMA *)
  // as ST:
  //   M_SENSOR_CIMA := SENSOR_CIMA;

// Rung 47
  LD %I0.13
  ST %M14                 (* FALHA_ÂNGULO *)
  // as ST:
  //   FALHA_ÂNGULO := %I0.13;

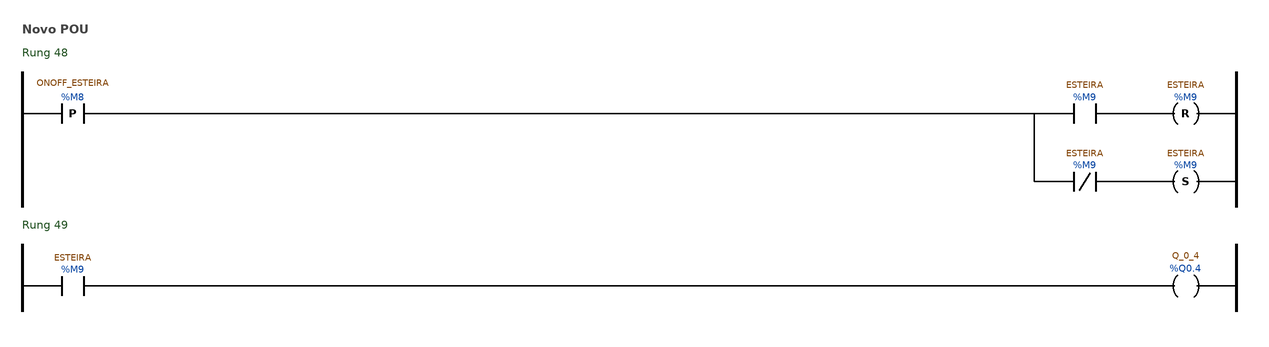

// Rung 48
  LDR %M8                 (* ONOFF_ESTEIRA *)
  MPS
  AND %M9                 (* ESTEIRA *)
  R %M9                   (* ESTEIRA *)
  MPP
  ANDN %M9                (* ESTEIRA *)
  S %M9                   (* ESTEIRA *)
  // as ST:
  //   IF RISING(ONOFF_ESTEIRA) AND ESTEIRA THEN ESTEIRA := FALSE; END_IF;
  //   IF RISING(ONOFF_ESTEIRA) AND NOT ESTEIRA THEN ESTEIRA := TRUE; END_IF;

// Rung 49
  LD %M9                  (* ESTEIRA *)
  ST %Q0.4                (* Q_0_4 *)
  // as ST:
  //   Q_0_4 := ESTEIRA;
